Staubli VAL3: utImage.pjx

--- utImage.pjx ---
Parameters version=s8.8.3Cs9_BS1660 stackSize=5000 millimeterUnit=true
Program file=start.pgx
Program file=stop.pgx
Data file=utImage.dtx
Type name=utAppearance path=./utAppearance/utAppearance.pjx
Type name=utBorder path=./utBorder/utBorder.pjx
Type name=utCommon path=./utCommon/utCommon.pjx
Type name=utEvents path=./utEvents/utEvents.pjx
Type name=utData path=./utData/utData.pjx

--- utImage.dtx ---
public utAppearance Appearance
  [0]
    string sBackgroundColour
    bool bVisibility
public utBorder Border
  [0]
    string sBorderColour
    string sBorderStyle
    num nBorderWidth
public utCommon Common
  [0]
    string sSourceImage
    string sID
    string sClass
    string sPage
public utEvents Events
  [0]
    bool bClick
    bool bMouseDown
    bool bMouseUp
public utData Data
  [0]
    num nVal
    bool bStatus
    string sSourceImg1
    string sSourceImg2

--- start.pgx ---
program start()
begin
end

--- stop.pgx ---
program stop()
begin
end
